(* IEC 61131-3 sources: plc-vscode/tests/st/test-ready/trust-platform/manual-tests/smoke/src, 2 files *)

(* ---- Math.st ---- *)
NAMESPACE Demo.Math
FUNCTION AddOne : DINT
VAR_INPUT
    X : DINT;
END_VAR
AddOne := X + 1;
END_FUNCTION
END_NAMESPACE

(* ---- Main.st ---- *)
USING Demo.Math;

PROGRAM Main
VAR
    value : DINT;
    result : DINT;
    t : TIME;
END_VAR

value := 41;
result := AddOne(value);
t := T#1s;

END_PROGRAM
